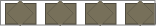
VISUALIZATION FRM_4InOutLed  // 156x26
VAR_IN_OUT    
    bLed1: BOOL;
    bLed2: BOOL;
    bLed3: BOOL;
    bLed4: BOOL;
    
   bLed1IsInput: BOOL;
   bLed2IsInput: BOOL;
   bLed3IsInput: BOOL;
   bLed4IsInput: BOOL;
END_VAR
    Rectangle (5,3 31x21), colour toggle: bLed1, invisible if: NOT bLed1IsInput
    Rectangle (45,3 31x21), colour toggle: bLed2, invisible if: NOT bLed2IsInput
    Rectangle (85,3 31x21), colour toggle: bLed3, invisible if: NOT bLed3IsInput
    Rectangle (125,3 31x21), colour toggle: bLed4, invisible if: NOT bLed4IsInput
    Polygon (7,13) (20,0) (33,13) (20,26) (20,26), colour toggle: bLed1, invisible if: bLed1IsInput
    Polygon (47,13) (60,0) (73,13) (60,26) (60,26), colour toggle: bLed2, invisible if: bLed2IsInput
    Polygon (87,13) (100,0) (113,13) (100,26) (100,26), colour toggle: bLed3, invisible if: bLed3IsInput
    Polygon (127,13) (140,0) (153,13) (140,26) (140,26), colour toggle: bLed4, invisible if: bLed4IsInput
END_VISUALIZATION

(* stored: Version 1.1.0.1
   Visu FRM_4InOutLed: Id {2599fefc-1291-0509-1a86-42db4f56ceb6} *)
